FUNCTION_BLOCK F (* Negative C4: two positions toggle, and each runs a copy of the CASE on the real position *)
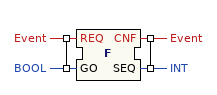
  EVENT_INPUT
    REQ WITH GO;
  END_EVENT
  EVENT_OUTPUT
    CNF WITH SEQ;
  END_EVENT
  VAR_INPUT
    GO : BOOL;
  END_VAR
  VAR_OUTPUT
    SEQ : INT;
  END_VAR
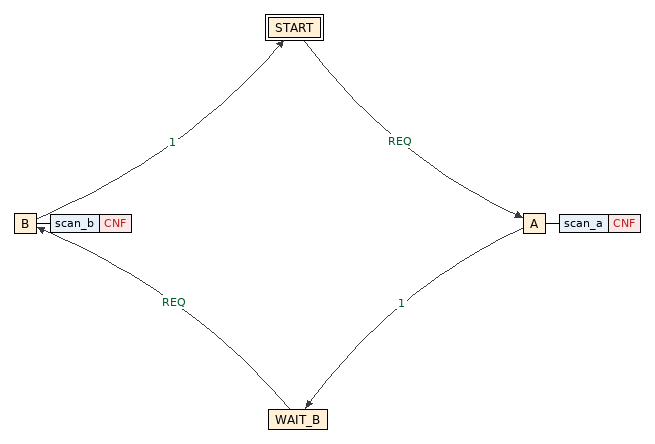
  EC_STATES
    START;
    A : scan_a -> CNF;
    WAIT_B;
    B : scan_b -> CNF;
  END_STATES
  EC_TRANSITIONS
    START TO A := REQ;
    A TO WAIT_B := 1;
    WAIT_B TO B := REQ;
    B TO START := 1;
  END_TRANSITIONS
  ALGORITHM scan_a IN ST:
CASE SEQ OF
  0:
    SEQ := 1;
  1:
    SEQ := 0;
END_CASE;
  END_ALGORITHM
  ALGORITHM scan_b IN ST:
CASE SEQ OF
  0:
    SEQ := 1;
  1:
    SEQ := 0;
END_CASE;
  END_ALGORITHM
END_FUNCTION_BLOCK
